(* IEC 61131-3 sources: plc-vscode/tests/st/test-ready/trust-platform/examples/ethercat_ek1100_elx008_v1/src, 2 files *)

(* ---- config.st ---- *)
CONFIGURATION Config
RESOURCE EtherCatRes ON PLC
    TASK MainTask (INTERVAL := T#10ms, PRIORITY := 1);
    PROGRAM P1 WITH MainTask : Main;
END_RESOURCE
VAR_CONFIG
    P1.DI0 AT %IX0.0 : BOOL;
    P1.DO0 AT %QX0.0 : BOOL;
END_VAR
END_CONFIGURATION

(* ---- Main.st ---- *)
PROGRAM Main
VAR
    RisingSeen : BOOL := FALSE;
    DI0 : BOOL;
    DO0 : BOOL;
END_VAR

IF DI0 THEN
    RisingSeen := TRUE;
END_IF;

DO0 := DI0 OR RisingSeen;
END_PROGRAM
